PROGRAM main
  VAR
    COLOR_SENSOR1 AT %QW1 : INT;
    COLOR_SENSOR2 AT %QW3 : INT;
    COLOR_SENSOR3 AT %QW5 : INT;
    DO_Conveyor AT %QX0.0 : BOOL;
    PUSHER1 AT %QX0.1 : BOOL;
    PUSHER2 AT %QX0.2 : BOOL;
    COUNT_RED AT %QX0.3 : BOOL;
    COUNT_YELLOW AT %QX0.4 : BOOL;
    COUNT_GREEN AT %QX0.5 : BOOL;
    COUNT_TOTAL AT %QX0.6 : BOOL;
    PB_START AT %QX0.7 : BOOL;
    PB_STOP_CONVEYOR AT %QX1.0 : BOOL;
    PB_STOP_RED AT %QX1.1 : BOOL;
    PB_STOP_YELLOW AT %QX1.2 : BOOL;
    PB_STOP_GREEN AT %QX1.3 : BOOL;
    PB_EMERGENCY AT %QX1.4 : BOOL;
    IS_RED : BOOL;
    IS_YELLOW : BOOL;
    IS_GREEN : BOOL;
    IS_ANY_BOX : BOOL;
    ENABLE_CONVEYOR : BOOL;
    ENABLE_RED : BOOL;
    ENABLE_YELLOW : BOOL;
    ENABLE_GREEN : BOOL;
    TP0 : TP;
    TP1 : TP;
    TP2 : TP;
  END_VAR

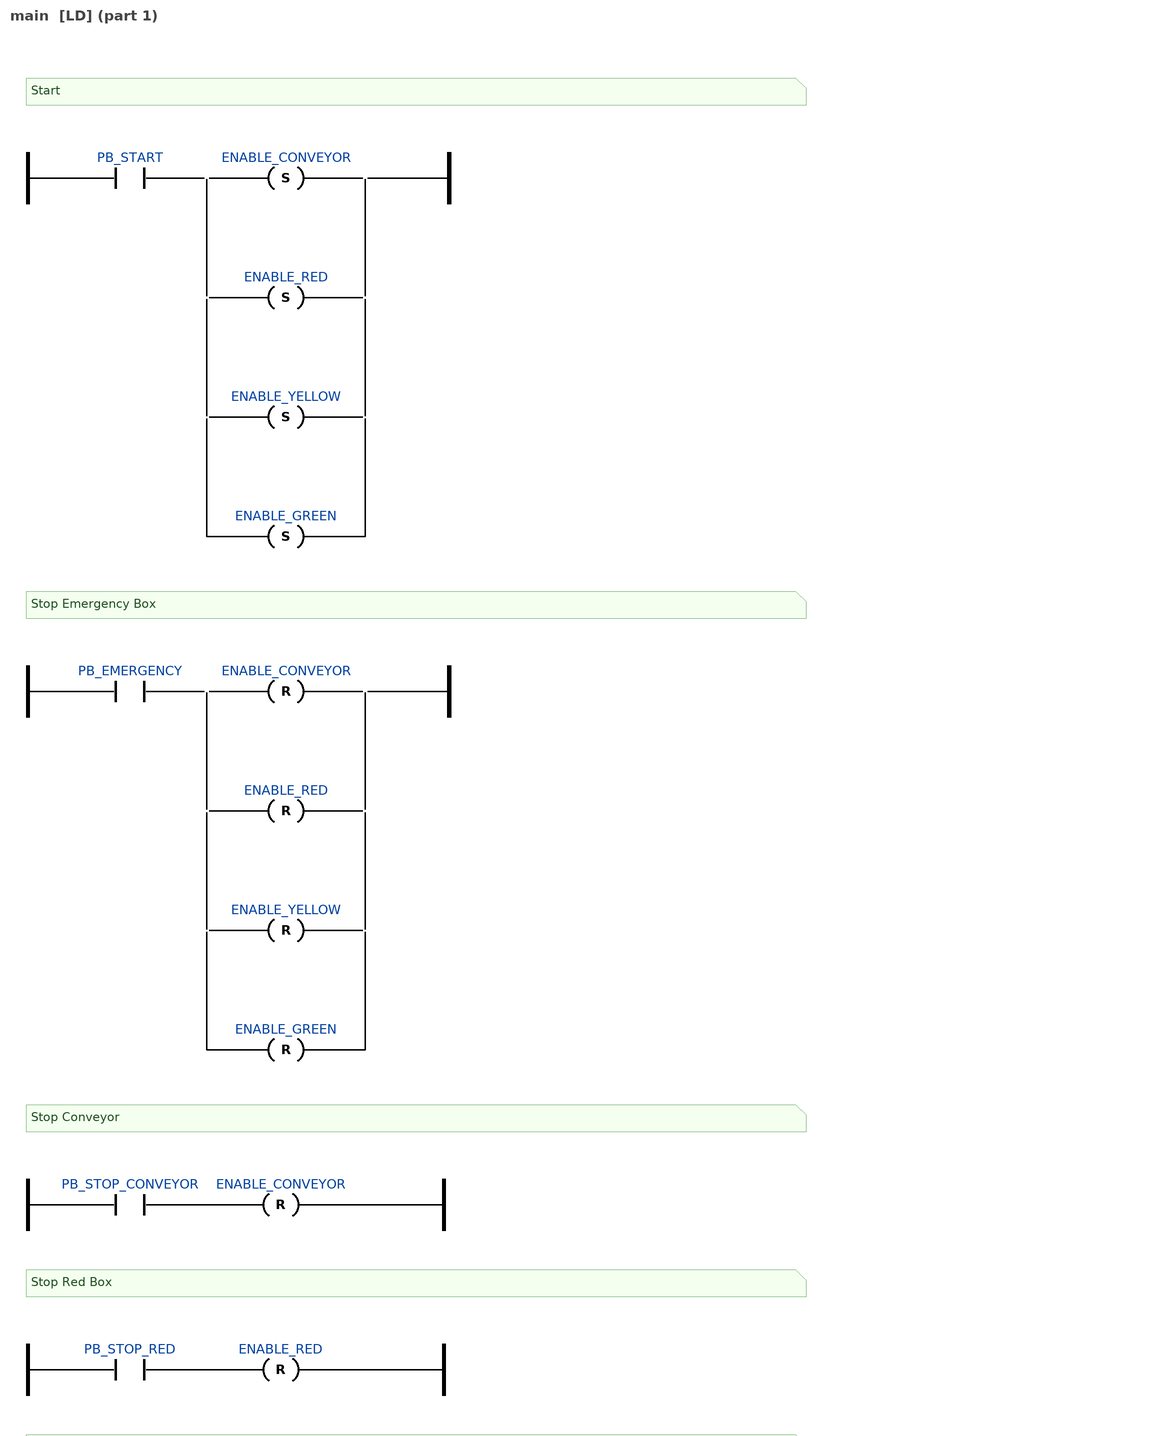
(* LD diagram, written out as Structured Text *)
(* Start *)
IF PB_START THEN ENABLE_CONVEYOR := TRUE; END_IF;
IF PB_START THEN ENABLE_RED := TRUE; END_IF;
IF PB_START THEN ENABLE_YELLOW := TRUE; END_IF;
IF PB_START THEN ENABLE_GREEN := TRUE; END_IF;
(* Stop Emergency Box *)
IF PB_EMERGENCY THEN ENABLE_CONVEYOR := FALSE; END_IF;
IF PB_EMERGENCY THEN ENABLE_RED := FALSE; END_IF;
IF PB_EMERGENCY THEN ENABLE_YELLOW := FALSE; END_IF;
IF PB_EMERGENCY THEN ENABLE_GREEN := FALSE; END_IF;
(* Stop Conveyor *)
IF PB_STOP_CONVEYOR THEN ENABLE_CONVEYOR := FALSE; END_IF;
(* Stop Red Box *)
IF PB_STOP_RED THEN ENABLE_RED := FALSE; END_IF;
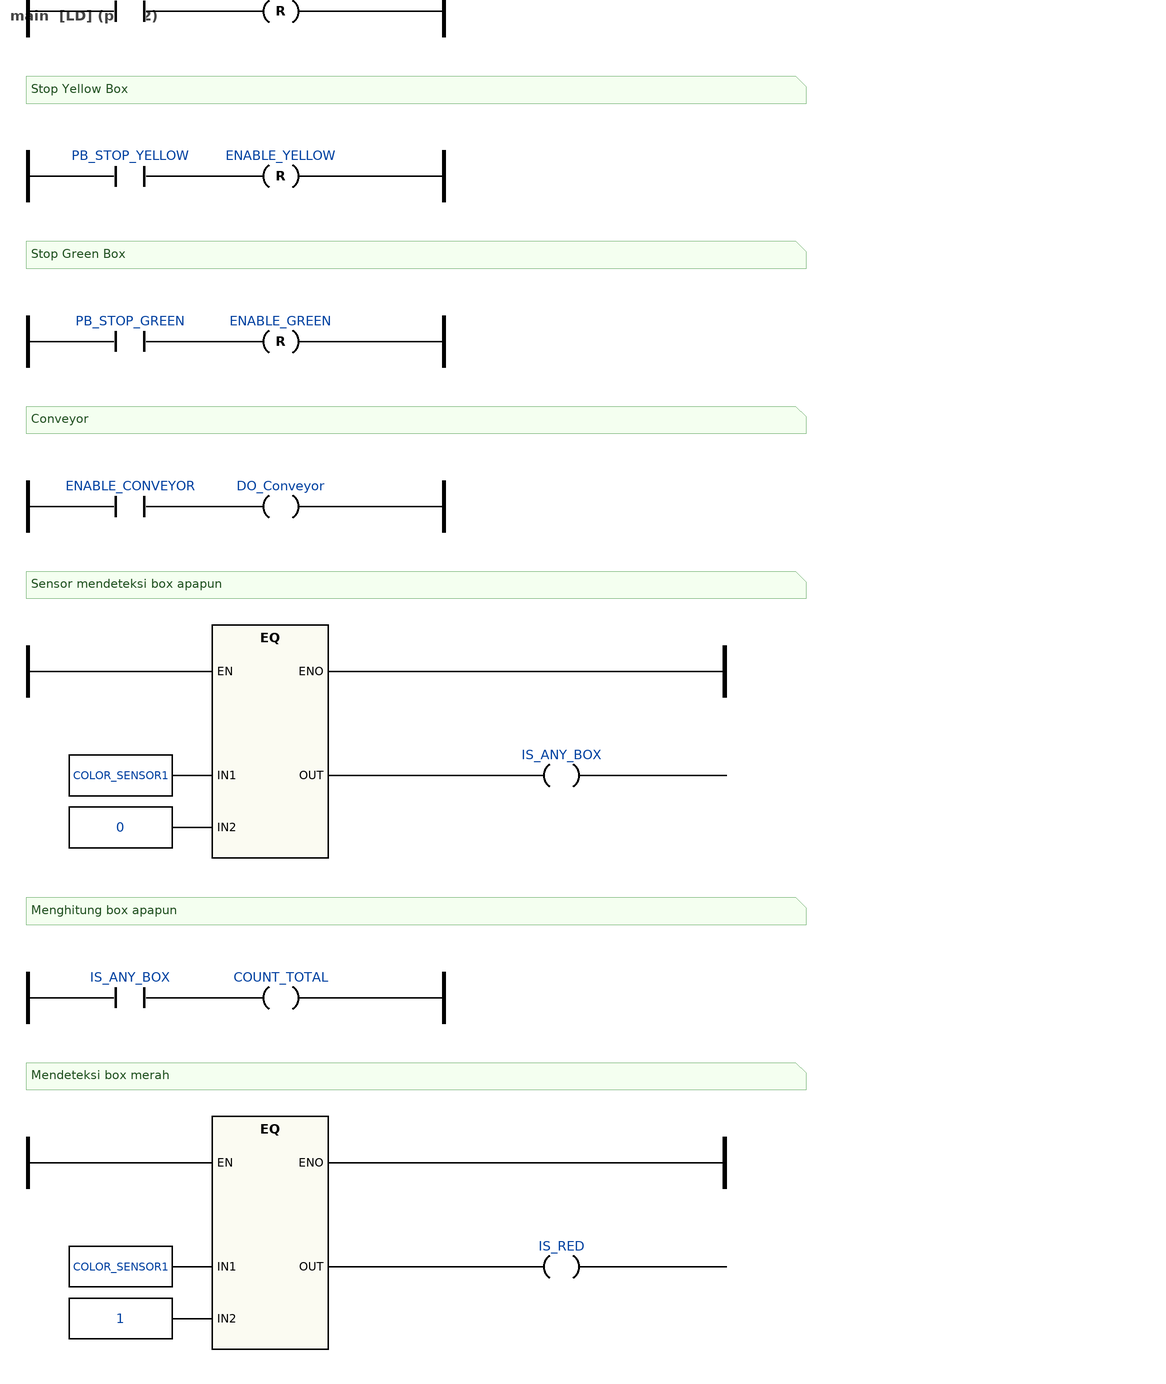
(* Stop Yellow Box *)
IF PB_STOP_YELLOW THEN ENABLE_YELLOW := FALSE; END_IF;
(* Stop Green Box *)
IF PB_STOP_GREEN THEN ENABLE_GREEN := FALSE; END_IF;
(* Conveyor *)
DO_Conveyor := ENABLE_CONVEYOR;
(* Sensor mendeteksi box apapun *)
IS_ANY_BOX := COLOR_SENSOR1 = 0;
(* Menghitung box apapun *)
COUNT_TOTAL := IS_ANY_BOX;
(* Mendeteksi box merah *)
IS_RED := COLOR_SENSOR1 = 1;
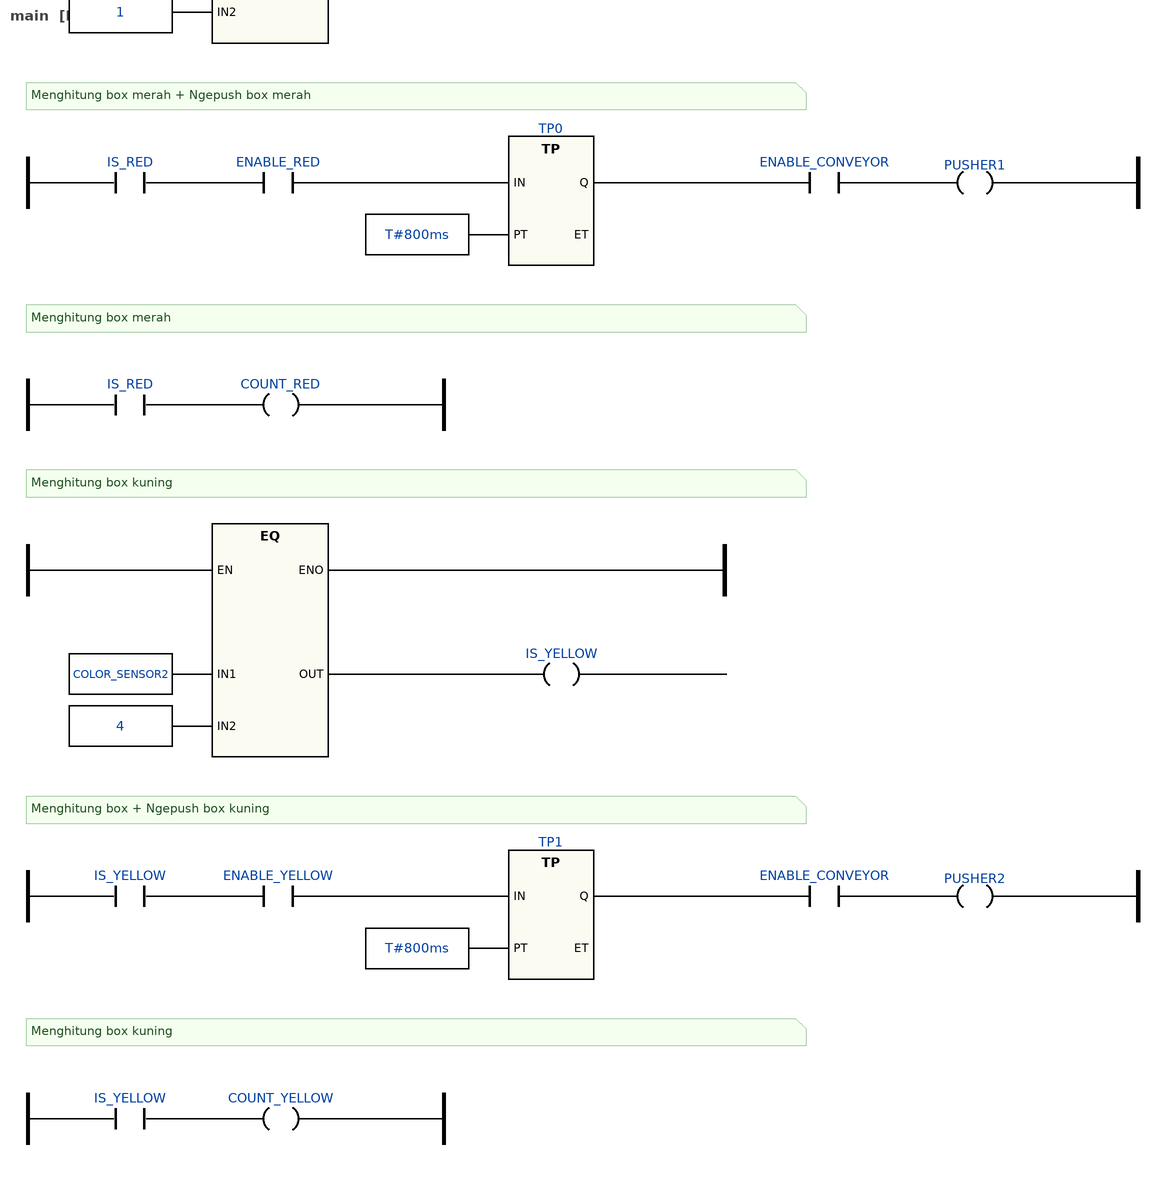
(* Menghitung box merah + Ngepush box merah *)
TP0(IN := IS_RED AND ENABLE_RED, PT := T#800ms);
PUSHER1 := TP0.Q AND ENABLE_CONVEYOR;
(* Menghitung box merah *)
COUNT_RED := IS_RED;
(* Menghitung box kuning *)
IS_YELLOW := COLOR_SENSOR2 = 4;
(* Menghitung box + Ngepush box kuning *)
TP1(IN := IS_YELLOW AND ENABLE_YELLOW, PT := T#800ms);
PUSHER2 := TP1.Q AND ENABLE_CONVEYOR;
(* Menghitung box kuning *)
COUNT_YELLOW := IS_YELLOW;
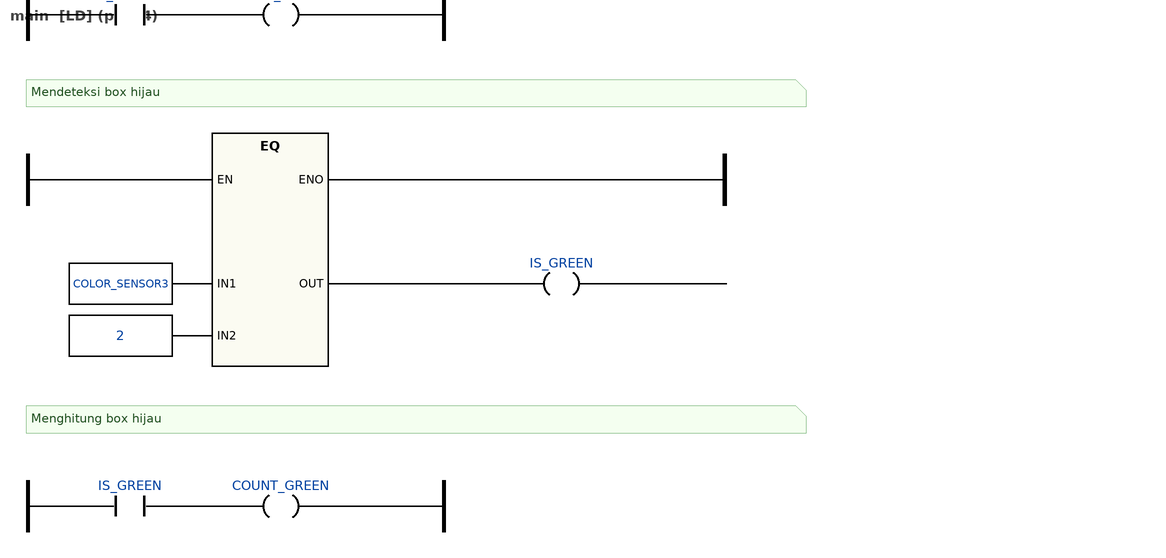
(* Mendeteksi box hijau *)
IS_GREEN := COLOR_SENSOR3 = 2;
(* Menghitung box hijau *)
COUNT_GREEN := IS_GREEN;
END_PROGRAM
